FUNCTION "F_AccessBenchProvision" : Void
{ S7_Optimized_Access := 'TRUE' }
VERSION : 0.1
BEGIN
        "FRK_LocalUsers".Count := 2;
        "FRK_LocalUsers".Rows[1].User := 'operator';
        "FRK_LocalUsers".Rows[1].Level := 1;
        "FRK_LocalUsers".Rows[1].Salt[0] := BYTE#16#A6;
        "FRK_LocalUsers".Rows[1].Salt[1] := BYTE#16#7F;
        "FRK_LocalUsers".Rows[1].Salt[2] := BYTE#16#A7;
        "FRK_LocalUsers".Rows[1].Salt[3] := BYTE#16#76;
        "FRK_LocalUsers".Rows[1].Salt[4] := BYTE#16#55;
        "FRK_LocalUsers".Rows[1].Salt[5] := BYTE#16#FA;
        "FRK_LocalUsers".Rows[1].Salt[6] := BYTE#16#32;
        "FRK_LocalUsers".Rows[1].Salt[7] := BYTE#16#65;
        "FRK_LocalUsers".Rows[1].Salt[8] := BYTE#16#ED;
        "FRK_LocalUsers".Rows[1].Salt[9] := BYTE#16#C7;
        "FRK_LocalUsers".Rows[1].Salt[10] := BYTE#16#41;
        "FRK_LocalUsers".Rows[1].Salt[11] := BYTE#16#31;
        "FRK_LocalUsers".Rows[1].Salt[12] := BYTE#16#C4;
        "FRK_LocalUsers".Rows[1].Salt[13] := BYTE#16#25;
        "FRK_LocalUsers".Rows[1].Salt[14] := BYTE#16#66;
        "FRK_LocalUsers".Rows[1].Salt[15] := BYTE#16#9C;
        "FRK_LocalUsers".Rows[1].PinHash[0] := BYTE#16#29;
        "FRK_LocalUsers".Rows[1].PinHash[1] := BYTE#16#11;
        "FRK_LocalUsers".Rows[1].PinHash[2] := BYTE#16#D1;
        "FRK_LocalUsers".Rows[1].PinHash[3] := BYTE#16#1F;
        "FRK_LocalUsers".Rows[1].PinHash[4] := BYTE#16#DD;
        "FRK_LocalUsers".Rows[1].PinHash[5] := BYTE#16#D0;
        "FRK_LocalUsers".Rows[1].PinHash[6] := BYTE#16#5A;
        "FRK_LocalUsers".Rows[1].PinHash[7] := BYTE#16#58;
        "FRK_LocalUsers".Rows[1].PinHash[8] := BYTE#16#01;
        "FRK_LocalUsers".Rows[1].PinHash[9] := BYTE#16#63;
        "FRK_LocalUsers".Rows[1].PinHash[10] := BYTE#16#2A;
        "FRK_LocalUsers".Rows[1].PinHash[11] := BYTE#16#D1;
        "FRK_LocalUsers".Rows[1].PinHash[12] := BYTE#16#74;
        "FRK_LocalUsers".Rows[1].PinHash[13] := BYTE#16#9A;
        "FRK_LocalUsers".Rows[1].PinHash[14] := BYTE#16#DB;
        "FRK_LocalUsers".Rows[1].PinHash[15] := BYTE#16#60;
        "FRK_LocalUsers".Rows[1].PinHash[16] := BYTE#16#25;
        "FRK_LocalUsers".Rows[1].PinHash[17] := BYTE#16#F6;
        "FRK_LocalUsers".Rows[1].PinHash[18] := BYTE#16#D8;
        "FRK_LocalUsers".Rows[1].PinHash[19] := BYTE#16#1B;
        "FRK_LocalUsers".Rows[1].PinHash[20] := BYTE#16#7A;
        "FRK_LocalUsers".Rows[1].PinHash[21] := BYTE#16#40;
        "FRK_LocalUsers".Rows[1].PinHash[22] := BYTE#16#BD;
        "FRK_LocalUsers".Rows[1].PinHash[23] := BYTE#16#DF;
        "FRK_LocalUsers".Rows[1].PinHash[24] := BYTE#16#AF;
        "FRK_LocalUsers".Rows[1].PinHash[25] := BYTE#16#F1;
        "FRK_LocalUsers".Rows[1].PinHash[26] := BYTE#16#80;
        "FRK_LocalUsers".Rows[1].PinHash[27] := BYTE#16#A9;
        "FRK_LocalUsers".Rows[1].PinHash[28] := BYTE#16#6E;
        "FRK_LocalUsers".Rows[1].PinHash[29] := BYTE#16#85;
        "FRK_LocalUsers".Rows[1].PinHash[30] := BYTE#16#0D;
        "FRK_LocalUsers".Rows[1].PinHash[31] := BYTE#16#87;
        "FRK_LocalUsers".Rows[2].User := 'admin';
        "FRK_LocalUsers".Rows[2].Level := 4;
        "FRK_LocalUsers".Rows[2].Salt[0] := BYTE#16#77;
        "FRK_LocalUsers".Rows[2].Salt[1] := BYTE#16#05;
        "FRK_LocalUsers".Rows[2].Salt[2] := BYTE#16#D0;
        "FRK_LocalUsers".Rows[2].Salt[3] := BYTE#16#D8;
        "FRK_LocalUsers".Rows[2].Salt[4] := BYTE#16#18;
        "FRK_LocalUsers".Rows[2].Salt[5] := BYTE#16#E9;
        "FRK_LocalUsers".Rows[2].Salt[6] := BYTE#16#72;
        "FRK_LocalUsers".Rows[2].Salt[7] := BYTE#16#4F;
        "FRK_LocalUsers".Rows[2].Salt[8] := BYTE#16#CC;
        "FRK_LocalUsers".Rows[2].Salt[9] := BYTE#16#34;
        "FRK_LocalUsers".Rows[2].Salt[10] := BYTE#16#18;
        "FRK_LocalUsers".Rows[2].Salt[11] := BYTE#16#20;
        "FRK_LocalUsers".Rows[2].Salt[12] := BYTE#16#95;
        "FRK_LocalUsers".Rows[2].Salt[13] := BYTE#16#7B;
        "FRK_LocalUsers".Rows[2].Salt[14] := BYTE#16#BB;
        "FRK_LocalUsers".Rows[2].Salt[15] := BYTE#16#4E;
        "FRK_LocalUsers".Rows[2].PinHash[0] := BYTE#16#53;
        "FRK_LocalUsers".Rows[2].PinHash[1] := BYTE#16#4C;
        "FRK_LocalUsers".Rows[2].PinHash[2] := BYTE#16#4C;
        "FRK_LocalUsers".Rows[2].PinHash[3] := BYTE#16#56;
        "FRK_LocalUsers".Rows[2].PinHash[4] := BYTE#16#88;
        "FRK_LocalUsers".Rows[2].PinHash[5] := BYTE#16#AA;
        "FRK_LocalUsers".Rows[2].PinHash[6] := BYTE#16#A4;
        "FRK_LocalUsers".Rows[2].PinHash[7] := BYTE#16#B6;
        "FRK_LocalUsers".Rows[2].PinHash[8] := BYTE#16#D9;
        "FRK_LocalUsers".Rows[2].PinHash[9] := BYTE#16#53;
        "FRK_LocalUsers".Rows[2].PinHash[10] := BYTE#16#10;
        "FRK_LocalUsers".Rows[2].PinHash[11] := BYTE#16#9E;
        "FRK_LocalUsers".Rows[2].PinHash[12] := BYTE#16#BC;
        "FRK_LocalUsers".Rows[2].PinHash[13] := BYTE#16#00;
        "FRK_LocalUsers".Rows[2].PinHash[14] := BYTE#16#15;
        "FRK_LocalUsers".Rows[2].PinHash[15] := BYTE#16#9B;
        "FRK_LocalUsers".Rows[2].PinHash[16] := BYTE#16#E1;
        "FRK_LocalUsers".Rows[2].PinHash[17] := BYTE#16#5A;
        "FRK_LocalUsers".Rows[2].PinHash[18] := BYTE#16#6A;
        "FRK_LocalUsers".Rows[2].PinHash[19] := BYTE#16#4D;
        "FRK_LocalUsers".Rows[2].PinHash[20] := BYTE#16#01;
        "FRK_LocalUsers".Rows[2].PinHash[21] := BYTE#16#8D;
        "FRK_LocalUsers".Rows[2].PinHash[22] := BYTE#16#C4;
        "FRK_LocalUsers".Rows[2].PinHash[23] := BYTE#16#13;
        "FRK_LocalUsers".Rows[2].PinHash[24] := BYTE#16#8A;
        "FRK_LocalUsers".Rows[2].PinHash[25] := BYTE#16#13;
        "FRK_LocalUsers".Rows[2].PinHash[26] := BYTE#16#2F;
        "FRK_LocalUsers".Rows[2].PinHash[27] := BYTE#16#9F;
        "FRK_LocalUsers".Rows[2].PinHash[28] := BYTE#16#6A;
        "FRK_LocalUsers".Rows[2].PinHash[29] := BYTE#16#96;
        "FRK_LocalUsers".Rows[2].PinHash[30] := BYTE#16#30;
        "FRK_LocalUsers".Rows[2].PinHash[31] := BYTE#16#95;

    "GDB_AccessPersistTest".ProvisionCount := "GDB_AccessPersistTest".ProvisionCount + 1;
    "StationA".Cell.Clamp.ParCfg.Timeout := T#30s;
    "StationA".Cell.Gate.ParCfg.Timeout := T#45s;
END_FUNCTION
FUNCTION "F_ConfigBenchPrepare" : Void
{ S7_Optimized_Access := 'TRUE' }
VERSION : 0.1
VAR_INPUT
    Startup : Bool;
END_VAR
VAR_TEMP
    StartupStamp : DTL;
    ResultCode : Int;
    SlotIndex : Int;
    Taken : Int;
    Accepted : Bool;
END_VAR
BEGIN
    "F_AlarmRecoveryDamage"(Startup := #Startup);
    IF #Startup THEN
        "StationA".Access.Policy.Required[11] := 3;
        "StationB".Access.Policy.Required[11] := 3;
    END_IF;
    IF #Startup THEN
        IF NOT "FRK_AccessStorage".UsersCommissioned AND "FRK_LocalUsers".SchemaVersion = 0 AND "FRK_LocalUsers".Generation = 0 AND "FRK_LocalUsers".Checksum = DWORD#0 THEN
            "F_AccessBenchProvision"();
        END_IF;
        "StationA".Access.Policy.Required[2] := 1;
        "StationA".Access.Policy.Required[4] := 1;
        "StationA".Access.Policy.Required[5] := 1;
        "StationA".Access.Policy.Required[8] := 4;
        "StationA".Access.Policy.SessionTimeout := T#0ms;
        "StationB".Access.Policy.Required[2] := 1;
        "StationB".Access.Policy.Required[4] := 1;
        "StationB".Access.Policy.Required[5] := 1;
        "StationB".Access.Policy.Required[8] := 4;
        "StationB".Access.Policy.SessionTimeout := T#0ms;
        "GDB_AccessTest".HashData[0] := BYTE#16#00;
        "GDB_AccessTest".HashData[1] := BYTE#16#01;
        "GDB_AccessTest".HashData[2] := BYTE#16#02;
        "GDB_AccessTest".HashData[3] := BYTE#16#03;
        "GDB_AccessTest".HashData[4] := BYTE#16#04;
        "GDB_AccessTest".HashData[5] := BYTE#16#05;
        "GDB_AccessTest".HashData[6] := BYTE#16#06;
        "GDB_AccessTest".HashData[7] := BYTE#16#07;
        "GDB_AccessTest".HashData[8] := BYTE#16#08;
        "GDB_AccessTest".HashData[9] := BYTE#16#09;
        "GDB_AccessTest".HashData[10] := BYTE#16#0A;
        "GDB_AccessTest".HashData[11] := BYTE#16#0B;
        "GDB_AccessTest".HashData[12] := BYTE#16#0C;
        "GDB_AccessTest".HashData[13] := BYTE#16#0D;
        "GDB_AccessTest".HashData[14] := BYTE#16#0E;
        "GDB_AccessTest".HashData[15] := BYTE#16#0F;
        "GDB_AccessTest".HashData[16] := BYTE#16#10;
        "GDB_AccessTest".HashData[17] := BYTE#16#11;
        "GDB_AccessTest".HashData[18] := BYTE#16#12;
        "GDB_AccessTest".HashData[19] := BYTE#16#13;
        "GDB_AccessTest".HashData[20] := BYTE#16#14;
        "GDB_AccessTest".HashData[21] := BYTE#16#15;
        "GDB_AccessTest".HashData[22] := BYTE#16#16;
        "GDB_AccessTest".HashData[23] := BYTE#16#17;
        "GDB_AccessTest".HashData[24] := BYTE#16#18;
        "GDB_AccessTest".HashData[25] := BYTE#16#19;
        "GDB_AccessTest".HashData[26] := BYTE#16#1A;
        "GDB_AccessTest".HashData[27] := BYTE#16#1B;
        "GDB_AccessTest".HashData[28] := BYTE#16#1C;
        "GDB_AccessTest".HashData[29] := BYTE#16#1D;
        "GDB_AccessTest".HashData[30] := BYTE#16#1E;
        "GDB_AccessTest".HashData[31] := BYTE#16#1F;
        "GDB_AccessTest".HashData[32] := BYTE#16#20;
        "GDB_AccessTest".HashData[33] := BYTE#16#21;
        "GDB_AccessTest".HashData[34] := BYTE#16#22;
        "GDB_AccessTest".HashData[35] := BYTE#16#23;
        "GDB_AccessTest".HashData[36] := BYTE#16#24;
        "GDB_AccessTest".HashData[37] := BYTE#16#25;
        "GDB_AccessTest".HashData[38] := BYTE#16#26;
        "GDB_AccessTest".HashData[39] := BYTE#16#27;
        "GDB_AccessTest".HashData[40] := BYTE#16#28;
        "GDB_AccessTest".HashData[41] := BYTE#16#29;
        "GDB_AccessTest".HashData[42] := BYTE#16#2A;
        "GDB_AccessTest".HashData[43] := BYTE#16#2B;
        "GDB_AccessTest".HashData[44] := BYTE#16#2C;
        "GDB_AccessTest".HashData[45] := BYTE#16#2D;
        "GDB_AccessTest".HashData[46] := BYTE#16#2E;
        "GDB_AccessTest".HashData[47] := BYTE#16#2F;
        "GDB_AccessTest".HashOk := "FRK_Sha256Pin"(Data := "GDB_AccessTest".HashData, Size := 0, Digest := "GDB_AccessTest".Hash0);
        "GDB_AccessTest".HashData[0] := BYTE#16#61;
        "GDB_AccessTest".HashData[1] := BYTE#16#62;
        "GDB_AccessTest".HashData[2] := BYTE#16#63;
        "GDB_AccessTest".HashData[3] := BYTE#16#00;
        "GDB_AccessTest".HashData[4] := BYTE#16#00;
        "GDB_AccessTest".HashData[5] := BYTE#16#00;
        "GDB_AccessTest".HashData[6] := BYTE#16#00;
        "GDB_AccessTest".HashData[7] := BYTE#16#00;
        "GDB_AccessTest".HashData[8] := BYTE#16#00;
        "GDB_AccessTest".HashData[9] := BYTE#16#00;
        "GDB_AccessTest".HashData[10] := BYTE#16#00;
        "GDB_AccessTest".HashData[11] := BYTE#16#00;
        "GDB_AccessTest".HashData[12] := BYTE#16#00;
        "GDB_AccessTest".HashData[13] := BYTE#16#00;
        "GDB_AccessTest".HashData[14] := BYTE#16#00;
        "GDB_AccessTest".HashData[15] := BYTE#16#00;
        "GDB_AccessTest".HashData[16] := BYTE#16#00;
        "GDB_AccessTest".HashData[17] := BYTE#16#00;
        "GDB_AccessTest".HashData[18] := BYTE#16#00;
        "GDB_AccessTest".HashData[19] := BYTE#16#00;
        "GDB_AccessTest".HashData[20] := BYTE#16#00;
        "GDB_AccessTest".HashData[21] := BYTE#16#00;
        "GDB_AccessTest".HashData[22] := BYTE#16#00;
        "GDB_AccessTest".HashData[23] := BYTE#16#00;
        "GDB_AccessTest".HashData[24] := BYTE#16#00;
        "GDB_AccessTest".HashData[25] := BYTE#16#00;
        "GDB_AccessTest".HashData[26] := BYTE#16#00;
        "GDB_AccessTest".HashData[27] := BYTE#16#00;
        "GDB_AccessTest".HashData[28] := BYTE#16#00;
        "GDB_AccessTest".HashData[29] := BYTE#16#00;
        "GDB_AccessTest".HashData[30] := BYTE#16#00;
        "GDB_AccessTest".HashData[31] := BYTE#16#00;
        "GDB_AccessTest".HashData[32] := BYTE#16#00;
        "GDB_AccessTest".HashData[33] := BYTE#16#00;
        "GDB_AccessTest".HashData[34] := BYTE#16#00;
        "GDB_AccessTest".HashData[35] := BYTE#16#00;
        "GDB_AccessTest".HashData[36] := BYTE#16#00;
        "GDB_AccessTest".HashData[37] := BYTE#16#00;
        "GDB_AccessTest".HashData[38] := BYTE#16#00;
        "GDB_AccessTest".HashData[39] := BYTE#16#00;
        "GDB_AccessTest".HashData[40] := BYTE#16#00;
        "GDB_AccessTest".HashData[41] := BYTE#16#00;
        "GDB_AccessTest".HashData[42] := BYTE#16#00;
        "GDB_AccessTest".HashData[43] := BYTE#16#00;
        "GDB_AccessTest".HashData[44] := BYTE#16#00;
        "GDB_AccessTest".HashData[45] := BYTE#16#00;
        "GDB_AccessTest".HashData[46] := BYTE#16#00;
        "GDB_AccessTest".HashData[47] := BYTE#16#00;
        "GDB_AccessTest".HashOk := "FRK_Sha256Pin"(Data := "GDB_AccessTest".HashData, Size := 3, Digest := "GDB_AccessTest".Hash1);
        "GDB_AccessTest".HashData[0] := BYTE#16#00;
        "GDB_AccessTest".HashData[1] := BYTE#16#01;
        "GDB_AccessTest".HashData[2] := BYTE#16#02;
        "GDB_AccessTest".HashData[3] := BYTE#16#03;
        "GDB_AccessTest".HashData[4] := BYTE#16#04;
        "GDB_AccessTest".HashData[5] := BYTE#16#05;
        "GDB_AccessTest".HashData[6] := BYTE#16#06;
        "GDB_AccessTest".HashData[7] := BYTE#16#07;
        "GDB_AccessTest".HashData[8] := BYTE#16#08;
        "GDB_AccessTest".HashData[9] := BYTE#16#09;
        "GDB_AccessTest".HashData[10] := BYTE#16#0A;
        "GDB_AccessTest".HashData[11] := BYTE#16#0B;
        "GDB_AccessTest".HashData[12] := BYTE#16#0C;
        "GDB_AccessTest".HashData[13] := BYTE#16#0D;
        "GDB_AccessTest".HashData[14] := BYTE#16#0E;
        "GDB_AccessTest".HashData[15] := BYTE#16#0F;
        "GDB_AccessTest".HashData[16] := BYTE#16#10;
        "GDB_AccessTest".HashData[17] := BYTE#16#11;
        "GDB_AccessTest".HashData[18] := BYTE#16#12;
        "GDB_AccessTest".HashData[19] := BYTE#16#13;
        "GDB_AccessTest".HashData[20] := BYTE#16#14;
        "GDB_AccessTest".HashData[21] := BYTE#16#15;
        "GDB_AccessTest".HashData[22] := BYTE#16#16;
        "GDB_AccessTest".HashData[23] := BYTE#16#17;
        "GDB_AccessTest".HashData[24] := BYTE#16#18;
        "GDB_AccessTest".HashData[25] := BYTE#16#19;
        "GDB_AccessTest".HashData[26] := BYTE#16#1A;
        "GDB_AccessTest".HashData[27] := BYTE#16#1B;
        "GDB_AccessTest".HashData[28] := BYTE#16#1C;
        "GDB_AccessTest".HashData[29] := BYTE#16#1D;
        "GDB_AccessTest".HashData[30] := BYTE#16#1E;
        "GDB_AccessTest".HashData[31] := BYTE#16#1F;
        "GDB_AccessTest".HashData[32] := BYTE#16#20;
        "GDB_AccessTest".HashData[33] := BYTE#16#21;
        "GDB_AccessTest".HashData[34] := BYTE#16#22;
        "GDB_AccessTest".HashData[35] := BYTE#16#23;
        "GDB_AccessTest".HashData[36] := BYTE#16#24;
        "GDB_AccessTest".HashData[37] := BYTE#16#25;
        "GDB_AccessTest".HashData[38] := BYTE#16#26;
        "GDB_AccessTest".HashData[39] := BYTE#16#27;
        "GDB_AccessTest".HashData[40] := BYTE#16#28;
        "GDB_AccessTest".HashData[41] := BYTE#16#29;
        "GDB_AccessTest".HashData[42] := BYTE#16#2A;
        "GDB_AccessTest".HashData[43] := BYTE#16#2B;
        "GDB_AccessTest".HashData[44] := BYTE#16#2C;
        "GDB_AccessTest".HashData[45] := BYTE#16#2D;
        "GDB_AccessTest".HashData[46] := BYTE#16#2E;
        "GDB_AccessTest".HashData[47] := BYTE#16#2F;
        "GDB_AccessTest".HashOk := "FRK_Sha256Pin"(Data := "GDB_AccessTest".HashData, Size := 32, Digest := "GDB_AccessTest".Hash2);
        "GDB_AccessTest".HashData[0] := BYTE#16#00;
        "GDB_AccessTest".HashData[1] := BYTE#16#01;
        "GDB_AccessTest".HashData[2] := BYTE#16#02;
        "GDB_AccessTest".HashData[3] := BYTE#16#03;
        "GDB_AccessTest".HashData[4] := BYTE#16#04;
        "GDB_AccessTest".HashData[5] := BYTE#16#05;
        "GDB_AccessTest".HashData[6] := BYTE#16#06;
        "GDB_AccessTest".HashData[7] := BYTE#16#07;
        "GDB_AccessTest".HashData[8] := BYTE#16#08;
        "GDB_AccessTest".HashData[9] := BYTE#16#09;
        "GDB_AccessTest".HashData[10] := BYTE#16#0A;
        "GDB_AccessTest".HashData[11] := BYTE#16#0B;
        "GDB_AccessTest".HashData[12] := BYTE#16#0C;
        "GDB_AccessTest".HashData[13] := BYTE#16#0D;
        "GDB_AccessTest".HashData[14] := BYTE#16#0E;
        "GDB_AccessTest".HashData[15] := BYTE#16#0F;
        "GDB_AccessTest".HashData[16] := BYTE#16#10;
        "GDB_AccessTest".HashData[17] := BYTE#16#11;
        "GDB_AccessTest".HashData[18] := BYTE#16#12;
        "GDB_AccessTest".HashData[19] := BYTE#16#13;
        "GDB_AccessTest".HashData[20] := BYTE#16#14;
        "GDB_AccessTest".HashData[21] := BYTE#16#15;
        "GDB_AccessTest".HashData[22] := BYTE#16#16;
        "GDB_AccessTest".HashData[23] := BYTE#16#17;
        "GDB_AccessTest".HashData[24] := BYTE#16#18;
        "GDB_AccessTest".HashData[25] := BYTE#16#19;
        "GDB_AccessTest".HashData[26] := BYTE#16#1A;
        "GDB_AccessTest".HashData[27] := BYTE#16#1B;
        "GDB_AccessTest".HashData[28] := BYTE#16#1C;
        "GDB_AccessTest".HashData[29] := BYTE#16#1D;
        "GDB_AccessTest".HashData[30] := BYTE#16#1E;
        "GDB_AccessTest".HashData[31] := BYTE#16#1F;
        "GDB_AccessTest".HashData[32] := BYTE#16#20;
        "GDB_AccessTest".HashData[33] := BYTE#16#21;
        "GDB_AccessTest".HashData[34] := BYTE#16#22;
        "GDB_AccessTest".HashData[35] := BYTE#16#23;
        "GDB_AccessTest".HashData[36] := BYTE#16#24;
        "GDB_AccessTest".HashData[37] := BYTE#16#25;
        "GDB_AccessTest".HashData[38] := BYTE#16#26;
        "GDB_AccessTest".HashData[39] := BYTE#16#27;
        "GDB_AccessTest".HashData[40] := BYTE#16#28;
        "GDB_AccessTest".HashData[41] := BYTE#16#29;
        "GDB_AccessTest".HashData[42] := BYTE#16#2A;
        "GDB_AccessTest".HashData[43] := BYTE#16#2B;
        "GDB_AccessTest".HashData[44] := BYTE#16#2C;
        "GDB_AccessTest".HashData[45] := BYTE#16#2D;
        "GDB_AccessTest".HashData[46] := BYTE#16#2E;
        "GDB_AccessTest".HashData[47] := BYTE#16#2F;
        "GDB_AccessTest".HashOk := "FRK_Sha256Pin"(Data := "GDB_AccessTest".HashData, Size := 48, Digest := "GDB_AccessTest".Hash3);
        "GDB_RoutingTest".PermitOne := TRUE;
        "GDB_RoutingTest".PermitTwo := TRUE;
        "GDB_RoutingTest".RootManualPermit := TRUE;
        "GDB_RoutingTest".NestedFinish := FALSE;
        "GDB_RoutingTest".InnerFinish := FALSE;
        "GDB_RoutingTest".NestedAccessLock := FALSE;
        #ResultCode := RD_SYS_T(OUT => #StartupStamp);
        IF #ResultCode = 0 THEN "GDB_UnitTest".BootStamp := DTL_TO_LDT(#StartupStamp); END_IF;
        "GDB_UnitTest".Restarts := "GDB_UnitTest".Restarts + 1;
        "GDB_UnitTest".FinishCycle := FALSE;
        "GDB_UnitTest".Permit := TRUE;
        "GDB_UnitTest".FaultRoot := FALSE;
        "GDB_UnitTest".ExitHold := FALSE;
        "GDB_UnitTest".IssueChild := FALSE;
        "GDB_UnitTest".LockStart := FALSE;
        "GDB_UnitTest".ChildCommand := 2;
        "GDB_UnitTest".Verdict := 1;
        "GDB_UnitTest".Reason := 2003;
        "GDB_UnitTest".CarrierControl := 0;
        "FRK_UnitSetLocalCarrier"(Unit := "StationA".Unit, Index := 1);
    END_IF;
    "GDB_FraktalHal".Data.StationA.Cell.Clamp.Finish := "GDB_UnitTest".FinishCycle;
    "GDB_FraktalHal".Data.StationA.Cell.Clamp.Permit := "GDB_UnitTest".Permit;
    "GDB_FraktalHal".Data.StationA.Cell.Clamp.ExitHold := "GDB_UnitTest".ExitHold;
    "GDB_FraktalHal".Data.StationA.Cell.Clamp.BackgroundFault := "GDB_UnitTest".FaultRoot;
    "GDB_FraktalHal".Data.StationA.Cell.Clamp.Verdict := "GDB_UnitTest".Verdict;
    "GDB_FraktalHal".Data.StationA.Cell.Clamp.Diag.ReasonCode := "GDB_UnitTest".Reason;
    "GDB_FraktalHal".Data.StationA.Cell.Clamp.Diag.Description := WSTRING#'test.start.permit';
    "GDB_FraktalHal".Data.StationA.Cell.Clamp.Diag.SourcePath := WSTRING#'StationA.Cell.Clamp';
    IF "GDB_UnitTest".IssueChild THEN
        "StationA".Cell.Clamp.Command := "GDB_UnitTest".ChildCommand;
        "StationA".Cell.Clamp.Execute := TRUE;
        "GDB_UnitTest".IssueChild := FALSE;
    END_IF;
    CASE "GDB_UnitTest".CarrierControl OF
        1: "FRK_UnitSetLocalCarrier"(Unit := "StationA".Unit, Index := 1);
        2: "FRK_Carriers".Slots[1].Enabled := FALSE;
        3: "FRK_Carriers".Slots[1].Context.Uid := 'other';
        ELSE "GDB_UnitTest".CarrierControl := 0;
    END_CASE;
    "GDB_UnitTest".CarrierControl := 0;
    "GDB_FraktalHal".Data.StationA.Cell.Gate.Permit := "GDB_RoutingTest".PermitOne;
    IF "GDB_RoutingTest".PermitTwo THEN "GDB_FraktalHal".Data.StationA.Cell.Gate.Sample := 0; ELSE "GDB_FraktalHal".Data.StationA.Cell.Gate.Sample := 1; END_IF;
    "GDB_FraktalHal".Data.StationA.Cell.Gate.Diag.ReasonCode := 2002;
    "GDB_FraktalHal".Data.StationA.Cell.Gate.Diag.Description := WSTRING#'test.manual.first';
    "GDB_FraktalHal".Data.StationA.Cell.Gate.LaterDiag.ReasonCode := 2003;
    "GDB_FraktalHal".Data.StationA.Cell.Gate.LaterDiag.Description := WSTRING#'test.manual.second';
    "GDB_FraktalHal".Data.StationA.Satellite.Cell.Clamp.Permit := "GDB_RoutingTest".RootManualPermit;
    "GDB_FraktalHal".Data.StationA.Satellite.Cell.Clamp.Diag.SourcePath := WSTRING#'StationA.Satellite.Cell.Clamp';
    "GDB_FraktalHal".Data.StationA.Satellite.Cell.Clamp.Diag.Description := WSTRING#'test.nested.permit';
    "GDB_FraktalHal".Data.StationA.Satellite.Cell.Clamp.Diag.ReasonCode := 2002;
    "GDB_FraktalHal".Data.StationA.Satellite.Inner.Cell.Clamp.Permit := TRUE;
    "GDB_FraktalHal".Data.StationA.Satellite.Cell.Clamp.Finish := "GDB_RoutingTest".NestedFinish;
    "GDB_FraktalHal".Data.StationA.Satellite.Inner.Cell.Clamp.Finish := "GDB_RoutingTest".InnerFinish;
    IF "GDB_RoutingTest".NestedAccessLock THEN
        "StationA".Satellite.Access.Policy.Required[5] := 4;
    ELSE
        "StationA".Satellite.Access.Policy.Required[5] := 0;
    END_IF;
    IF "GDB_RoutingTest".LocalPulse THEN
        "GDB_RoutingTest".LocalRequest.Kind := "GDB_RoutingTest".LocalKind;
        "GDB_RoutingTest".LocalRequest.IntValue := "GDB_RoutingTest".LocalValue;
        "FRK_UnitOperation"(Core := "StationA".Satellite.Core, Unit := "StationA".Satellite.Unit, Status := "StationA".Satellite.Status, Policy := "StationA".Satellite.ModePolicy, Access := "StationA".Satellite.Access, Supported := "StationA".Satellite.SupportedModesPublished, Request := "GDB_RoutingTest".LocalRequest, Response := "FRK_UnitScratch".Response, Trusted := FALSE);
        "GDB_RoutingTest".LocalAccepted := "FRK_UnitScratch".Response.Accepted;
        "GDB_RoutingTest".LocalFirstKind := -1;
        IF "FRK_UnitScratch".Response.Report.Count > 0 THEN "GDB_RoutingTest".LocalFirstKind := "FRK_UnitScratch".Response.Report.Reasons[1].Kind; END_IF;
        "GDB_RoutingTest".LocalPulse := FALSE;
    END_IF;
    "StationA".Access.ProviderEnabled := NOT "GDB_AccessTest".ProviderOff;
    "StationB".Access.ProviderEnabled := NOT "GDB_AccessTest".ProviderOff;
    "StationA".AlarmLog.SinkEnabled := TRUE;
    "StationB".AlarmLog.SinkEnabled := TRUE;
    "GDB_FraktalHal".Data.StationA.Cell.Clamp.Sample := "GDB_StateAlarmTest".Position;
    IF "GDB_StateAlarmTest".ClearLog THEN
        "FRK_AlarmBegin"(AlarmLog := "StationA".AlarmLog, Startup := TRUE);
        "GDB_StateAlarmTest".SinkCome := 0;
        "GDB_StateAlarmTest".SinkClose := 0;
        "GDB_StateAlarmTest".ClearLog := FALSE;
    END_IF;
    IF "GDB_StateAlarmTest".RaisePulse THEN
        "GDB_StateAlarmTest".Slot := "FRK_AlarmRaise"(AlarmLog := "StationA".AlarmLog, Diag := "GDB_StateAlarmTest".Diag, ResetClass := "GDB_StateAlarmTest".ResetClass);
        "GDB_StateAlarmTest".RaisePulse := FALSE;
    END_IF;
    IF "GDB_StateAlarmTest".GonePulse THEN
        "GDB_StateAlarmTest".GoneAccepted := "FRK_AlarmGone"(AlarmLog := "StationA".AlarmLog, Slot := "GDB_StateAlarmTest".Slot);
        "GDB_StateAlarmTest".GonePulse := FALSE;
    END_IF;
    IF "GDB_StateAlarmTest".FillPulse THEN
        FOR #SlotIndex := 1 TO "GDB_StateAlarmTest".FillCount DO
            #Taken := "FRK_AlarmRaise"(AlarmLog := "StationA".AlarmLog, Diag := "GDB_StateAlarmTest".Diag, ResetClass := "GDB_StateAlarmTest".ResetClass);
            IF "GDB_StateAlarmTest".ResetClass = 0 THEN #Accepted := "FRK_AlarmGone"(AlarmLog := "StationA".AlarmLog, Slot := #Taken); END_IF;
        END_FOR;
        "GDB_StateAlarmTest".FillPulse := FALSE;
    END_IF;
    IF "GDB_StateAlarmTest".CauseLive THEN
        IF "GDB_StateAlarmTest".CauseSlot = 0 THEN
            "GDB_StateAlarmTest".CauseSlot := "FRK_AlarmRaise"(AlarmLog := "StationA".AlarmLog, Diag := "GDB_StateAlarmTest".Diag, ResetClass := 1);
        ELSIF "StationA".AlarmLog.Active["GDB_StateAlarmTest".CauseSlot].State = 0 THEN
            "GDB_StateAlarmTest".CauseSlot := "FRK_AlarmRaise"(AlarmLog := "StationA".AlarmLog, Diag := "GDB_StateAlarmTest".Diag, ResetClass := 1);
        END_IF;
    ELSIF "GDB_StateAlarmTest".CauseSlot > 0 THEN
        #Accepted := "FRK_AlarmGone"(AlarmLog := "StationA".AlarmLog, Slot := "GDB_StateAlarmTest".CauseSlot);
        "GDB_StateAlarmTest".CauseSlot := 0;
    END_IF;
    "FRK_StateSweep"(Flags := "GDB_StateAlarmTest".StandaloneFlags, Count := "GDB_StateAlarmTest".StandaloneCount, Touched := "GDB_StateAlarmTest".Touched, Startup := #Startup);
    IF "GDB_StateAlarmTest".PublishState THEN
        "GDB_StateAlarmTest".StandaloneReturn := "FRK_State"(Idx := "GDB_StateAlarmTest".StateIndex, Key := 'project.state.atHome', Ok := "GDB_StateAlarmTest".StateValue, Flags := "GDB_StateAlarmTest".StandaloneFlags, Count := "GDB_StateAlarmTest".StandaloneCount, Touched := "GDB_StateAlarmTest".Touched);
    END_IF;
    "FRK_ConfigRuntime".Unavailable := "GDB_ConfigTest".Unavailable;
    IF "GDB_ConfigTest".BlockRestore THEN "StationA".ConfigPersist.RestorePolicy := 1;
    ELSE "StationA".ConfigPersist.RestorePolicy := 0; END_IF;
    IF "GDB_ConfigTest".CorruptPulse THEN
        "GDB_ConfigTest".CorruptSlot := "FRK_ConfigFind"(Scope := "GDB_ConfigTest".CorruptScope, Key := "GDB_ConfigTest".CorruptKey, ModelCode := "GDB_ConfigTest".CorruptModel);
        IF "GDB_ConfigTest".CorruptSlot > 0 THEN
            "FRK_ConfigStore".Rows["GDB_ConfigTest".CorruptSlot].SchemaVersion := "GDB_ConfigTest".CorruptSchema;
            "FRK_ConfigStore".Rows["GDB_ConfigTest".CorruptSlot].Record.ValueText := "GDB_ConfigTest".CorruptText;
        END_IF;
        "GDB_ConfigTest".CorruptPulse := FALSE;
    END_IF;
    "StationA".Cell.Clamp.ParCfg.Timeout := T#30s;
    "StationA".Cell.Gate.ParCfg.Timeout := T#45s;
END_FUNCTION

FUNCTION "F_ConfigBenchObserve" : Void
{ S7_Optimized_Access := 'TRUE' }
VERSION : 0.1
VAR_INPUT
    Startup : Bool;
END_VAR
BEGIN
    "GDB_StateAlarmTest".NativeFaultSlot := "StationA".Cell.Gate.Core.FaultSlot;
    "GDB_RoutingTest".ManExecute := "StationA".Cell.Gate.Execute;
    "GDB_RoutingTest".ManStarts := "StationA".Cell.Gate.Device.StartCount;
    "GDB_UnitTest".Scans := "GDB_UnitTest".Scans + 1;
    "GDB_UnitTest".ChildExecute := "StationA".Cell.Clamp.Execute;
    "GDB_UnitTest".ChildState := "StationA".Cell.Clamp.Core.Exec;
    "GDB_UnitTest".CarrierWrites := "FRK_Carriers".Slots[1].Writes;
    "GDB_UnitTest".CarrierSerial := "FRK_Carriers".Slots[1].Serial;
    "GDB_UnitTest".WrittenUid := "FRK_Carriers".Slots[1].Written.Uid;
    "GDB_UnitTest".WrittenVerdict := "FRK_Carriers".Slots[1].Written.Result.Verdict;
    IF "StationA".AlarmLog.RingHead > 0 AND "StationA".AlarmLog.RingHead <= 64 THEN
        "GDB_UnitTest".LastEvent := "StationA".AlarmLog.Ring["StationA".AlarmLog.RingHead].ReasonCode;
    END_IF;
    "GDB_UnitTest".SecretCleared := "StationA".HmiRequest.Secret = '';
    "GDB_UnitTest".SnapshotSecretCleared := "StationA".Unit.Request.Secret = '';
    IF "StationA".Access.LoginBusy AND ("GDB_AccessTest".CancelOnLogin OR "GDB_AccessTest".SupersedeOnLogin) THEN
        "GDB_AccessTest".InterruptedBusy := TRUE;
        IF "GDB_AccessTest".CancelOnLogin THEN
            "GDB_AccessTest".InterruptRequest.Kind := 2;
            "FRK_UnitOperation"(Core := "StationA".Core, Unit := "StationA".Unit, Status := "StationA".Status, Policy := "StationA".ModePolicy, Access := "StationA".Access, Supported := "StationA".SupportedModesPublished, Request := "GDB_AccessTest".InterruptRequest, Response := "FRK_UnitScratch".Response, Trusted := FALSE);
        ELSE
            "GDB_AccessTest".SupersededSequence := "FRK_AccessNext"(Previous := "StationA".Access.LoginSequence);
            "FRK_AccessLogin"(Access := "StationA".Access, User := 'unknown', Secret := 'wrong', Sequence := "GDB_AccessTest".SupersededSequence);
        END_IF;
        "GDB_AccessTest".CancelOnLogin := FALSE;
        "GDB_AccessTest".SupersedeOnLogin := FALSE;
    END_IF;
    "F_ConfigSetBench"();
    "F_AccessPersistenceBench"(Startup := #Startup);
    "F_AlarmPersistenceBench"();
    "F_AlarmRecoveryBench"();
    "F_TestSequenceQuiesce"();
END_FUNCTION
